(* IEC 61131-3 sources: PLC--Learning/exercises, 3 files *)

(* ---- 01_math_bool.st ---- *)
   // Exercise 01: Math + Boolean basics
   PROGRAM PLC_PRG
   VAR
       a       : INT := 5;
       b       : INT := 3;
       sum     : INT;
       product : INT;
       x       : BOOL;
       y       : BOOL;
       both    : BOOL;
       result  : BOOL;
   END_VAR

   sum     := a + b;
   product := a * b;
   both    := x AND y;
   result  := x XOR y;

(* ---- 02_math_compare.st ---- *)
// Exercise 02: Math (+ - * /) and comparisons with IF
// Note: INT division cuts off decimals (28/26 = 1)
PROGRAM Ex02_Compare
VAR
    // Math
    num1      : INT := 10;
    num2      : INT := 4;
    addResult : INT;
    subResult : INT;
    mulResult : INT;
    divResult : INT;

    // Temperature
    temp   : INT := 20;
    isHot  : BOOL;
    isCold : BOOL;
    fan    : BOOL;
    heater : BOOL;
END_VAR

// Math
addResult := num1 + num2;
subResult := num1 - num2;
mulResult := num1 * num2;
divResult := num1 / num2;

// Temperature checks
isHot  := temp > 30;
isCold := temp < 15;

// Decisions
IF isHot THEN
    fan := TRUE;
ELSE
    fan := FALSE;
END_IF

IF isCold THEN
    heater := TRUE;
ELSE
    heater := FALSE;
END_IF

(* ---- 03_real_or_not.st ---- *)
// Exercise 03: REAL numbers, OR, NOT
// REAL keeps decimals: 28.0 / 26.0 = 1.0769...
PROGRAM Ex03_Real
VAR
    // Decimals
    r1      : REAL := 28.0;
    r2      : REAL := 26.0;
    realDiv : REAL;
    average : REAL;

    // Machine safety
    doorOpen   : BOOL;
    emergency  : BOOL;
    alarm      : BOOL;
    doorClosed : BOOL;
    machineRun : BOOL;
END_VAR

// Decimals
realDiv := r1 / r2;
average := (r1 + r2) / 2.0;

// Machine safety
alarm      := doorOpen OR emergency;
doorClosed := NOT doorOpen;
machineRun := NOT alarm;
